// TIA Portal V20 export
Screen "160FX1Layout"  1276x673
  ScreenItem "Line_Header_X0_Y64" at 0,64 size 1276x0  Type=HmiLine
  ScreenItem "permanentareaborderrectangle" at 0,0 size 0x0  Type=HmiRectangle
  ScreenItem "Button_Back" at 2,2 size 90x60  Type=HmiButton
  ScreenItem "Fusszeile_Button_ManualOPMode1_2" at 279,2 size 90x60  Type=HmiButton
  ScreenItem "文本域_3" at 1107,71 size 139x22  Type=HmiTextBox
  ScreenItem "文本域_1" at 1107,160 size 156x23  Type=HmiTextBox
  ScreenItem "文本域_2" at 1107,246 size 135x23  Type=HmiTextBox
  ScreenItem "文本域_22" at 1124,402 size 104x23  Type=HmiTextBox
  ScreenItem "Fusszeile_Button_ManualOPMode1_1" at 95,2 size 90x60  Type=HmiButton
  ScreenItem "Button_Back_1" at 1180,606 size 90x60  Type=HmiButton
  ScreenItem "Fusszeile_Button_ManualOPMode1_3" at 187,2 size 90x60  Type=HmiButton
  ScreenItem "Fusszeile_Button_ManualOPMode1_4" at 997,2 size 90x60  Type=HmiButton
  ScreenItem "Fusszeile_Button_ManualOPMode1_5" at 902,1 size 90x60  Type=HmiButton
  ScreenItem "文本域_14" at 936,-172 size 140x40  Type=HmiTextBox
  ScreenItem "文本域_5" at -1,82 size 120x40  Type=HmiTextBox
  ScreenItem "Title_ScreenOverview_X390_Y2_1" at 384,5 size 510x57  Type=HmiTextBox
  ScreenItem "文本域_27" at -1,126 size 120x40  Type=HmiTextBox
  ScreenItem "Graphic view_1" at 19,230 size 860x259  Type=HmiGraphicView
  ScreenItem "Line_9" at 558,162 size 94x182  Type=HmiLine
  ScreenItem "Line_2" at 702,237 size 20x91  Type=HmiLine
  ScreenItem "Line_5" at 752,186 size 92x151  Type=HmiLine
  ScreenItem "Line_17" at 108,206 size 171x117  Type=HmiLine
  ScreenItem "Line_6" at 751,373 size 177x7  Type=HmiLine
  ScreenItem "Line_10" at 514,412 size 202x102  Type=HmiLine
  ScreenItem "Line_13" at 646,414 size 83x147  Type=HmiLine
  ScreenItem "Line_1" at 375,375 size 288x138  Type=HmiLine
  ScreenItem "Line_18" at 217,417 size 62x96  Type=HmiLine
  ScreenItem "Line_16" at 79,341 size 76x150  Type=HmiLine
  ScreenItem "文本域_6" at 11,477 size 140x40  Type=HmiTextBox
  ScreenItem "文本域_7" at 168,516 size 100x20  Type=HmiTextBox
  ScreenItem "文本域_8" at 321,510 size 100x40  Type=HmiTextBox
  ScreenItem "文本域_9" at 455,517 size 100x20  Type=HmiTextBox
  ScreenItem "文本域_10" at 565,533 size 140x40  Type=HmiTextBox
  ScreenItem "文本域_12" at 921,359 size 100x40  Type=HmiTextBox
  ScreenItem "文本域_13" at 502,110 size 140x20  Type=HmiTextBox
  ScreenItem "文本域_15" at 921,192 size 140x40  Type=HmiTextBox
  ScreenItem "文本域_17" at 18,170 size 100x20  Type=HmiTextBox
  ScreenItem "文本域_18" at 652,176 size 100x20  Type=HmiTextBox
  ScreenItem "文本域_20" at 766,130 size 140x20  Type=HmiTextBox
  ScreenItem "文本域_21" at 128,98 size 140x40  Type=HmiTextBox
  ScreenItem "文本域_23" at 281,98 size 140x40  Type=HmiTextBox
  ScreenItem "Line_11" at 347,179 size 75x122  Type=HmiLine
  ScreenItem "Line_4" at 190,174 size 228x146  Type=HmiLine
  ScreenItem "Line_12" at 777,224 size 144x115  Type=HmiLine
  ScreenItem "Line_19" at 777,402 size 186x161  Type=HmiLine
  ScreenItem "文本域_26" at 907,533 size 140x40  Type=HmiTextBox
  ScreenItem "文本域_4" at 753,526 size 140x20  Type=HmiTextBox
  ScreenItem "Line_3" at 753,409 size 37x112  Type=HmiLine
  ScreenItem "Faceplate container_5" at 36,189 size 59x45  Type=HmiFaceplateContainer
  ScreenItem "面板容器_10" at 502,131 size 153x58  Type=HmiFaceplateContainer
  ScreenItem "Faceplate container_1" at 670,197 size 59x45  Type=HmiFaceplateContainer
  ScreenItem "面板容器_7" at 761,151 size 148x58  Type=HmiFaceplateContainer
  ScreenItem "面板容器_6" at 921,233 size 149x54  Type=HmiFaceplateContainer
  ScreenItem "Faceplate container_4" at 941,399 size 59x45  Type=HmiFaceplateContainer
  ScreenItem "面板容器_15" at 907,573 size 149x54  Type=HmiFaceplateContainer
  ScreenItem "面板容器_9" at 753,547 size 148x58  Type=HmiFaceplateContainer
  ScreenItem "面板容器_20" at 565,573 size 150x51  Type=HmiFaceplateContainer
  ScreenItem "面板容器_4" at 477,540 size 56x46  Type=HmiFaceplateContainer
  ScreenItem "Faceplate container_2" at 187,539 size 61x45  Type=HmiFaceplateContainer
  ScreenItem "面板容器_5" at 11,518 size 143x50  Type=HmiFaceplateContainer
  ScreenItem "Faceplate container_3" at 341,550 size 59x45  Type=HmiFaceplateContainer
  ScreenItem "LSicar_Valve8Pos_LeftHomeRightWork_WithPB_5" at 1099,95 size 160x53  Type=HmiFaceplateContainer
  ScreenItem "LSicar_Valve8Pos_LeftHomeRightWork_WithPB_1" at 1099,183 size 160x53  Type=HmiFaceplateContainer
  ScreenItem "LSicar_Valve8Pos_LeftHomeRightWork_WithPB_2" at 1099,269 size 160x53  Type=HmiFaceplateContainer
  ScreenItem "面板容器_22" at 1061,435 size 96x32  Type=HmiFaceplateContainer
  ScreenItem "面板容器_23" at 1171,435 size 96x32  Type=HmiFaceplateContainer
  ScreenItem "Move_Legend" at 1182,2 size 90x60  Type=HmiButton
  ScreenItem "面板容器_2" at 1090,4 size 88x58  Type=HmiFaceplateContainer
  ScreenItem "OPMode1_Blocked" at 1164,6 size 14x14  Type=HmiGraphicView
  ScreenItem "OPMode4_Foreground_Blocked" at 1091,4 size 88x58  Type=HmiGraphicView
  ScreenItem "Button_Back_3" at 122,606 size 90x60  Type=HmiButton
  ScreenItem "Button_Back_2" at 8,606 size 90x60  Type=HmiButton
  ScreenItem "面板容器_11" at 282,137 size 150x51  Type=HmiFaceplateContainer
  ScreenItem "面板容器_8" at 130,139 size 144x51  Type=HmiFaceplateContainer
